(* IEC 61131-3 sources: llm-plc-st-eval/data/definitivo/claude-sonnet-4-6/B2/zero_shot, 3 files *)

(* ---- ejec_1.st ---- *)
```pascal
FUNCTION_BLOCK FB_Valvula
VAR_INPUT
    nivelAlto : BOOL; (* Sensor de nivel alto del tanque *)
END_VAR

VAR_OUTPUT
    valvula : BOOL; (* TRUE = válvula abierta, FALSE = válvula cerrada *)
END_VAR

VAR
    tonRetardo : TON; (* Temporizador de retardo para confirmación de nivel alto *)
END_VAR

(*
    Control de válvula de drenaje:
    - La válvula abre cuando nivelAlto permanece activo durante 5 segundos continuos.
    - La válvula cierra de inmediato si nivelAlto deja de estar activo.
*)

(* Activar temporizador solo mientras nivelAlto esté activo *)
tonRetardo(IN := nivelAlto, PT := T#5S);

(* La válvula abre cuando el temporizador completa los 5 segundos *)
(* Si nivelAlto cae, tonRetardo.Q se resetea de inmediato y la válvula cierra *)
valvula := tonRetardo.Q;

END_FUNCTION_BLOCK
```

(* ---- ejec_2.st ---- *)
```pascal
FUNCTION_BLOCK FB_Valvula
VAR_INPUT
    nivelAlto : BOOL; (* Sensor de nivel alto del tanque *)
END_VAR

VAR_OUTPUT
    valvula : BOOL; (* TRUE = válvula abierta, FALSE = válvula cerrada *)
END_VAR

VAR
    tonRetardo : TON; (* Temporizador de retardo para confirmar nivel alto *)
END_VAR

(*
    Control de válvula de drenaje:
    - La válvula abre cuando nivelAlto permanece activo durante 5 segundos continuos.
    - La válvula cierra de inmediato si nivelAlto deja de estar activo.
*)

(* Activar temporizador solo mientras nivelAlto esté activo *)
tonRetardo(IN := nivelAlto, PT := T#5S);

(* La válvula abre cuando el temporizador completa los 5 segundos *)
(* Si nivelAlto cae, tonRetardo.Q se pone FALSE de inmediato (IN=FALSE resetea el TON) *)
valvula := tonRetardo.Q;

END_FUNCTION_BLOCK
```

(* ---- ejec_3.st ---- *)
```pascal
FUNCTION_BLOCK FB_Valvula
VAR_INPUT
    nivelAlto : BOOL; (* Sensor de nivel alto del tanque *)
END_VAR

VAR_OUTPUT
    valvula : BOOL; (* TRUE = válvula abierta, FALSE = válvula cerrada *)
END_VAR

VAR
    tonRetardo : TON; (* Temporizador de retardo para confirmar nivel alto *)
END_VAR

(* ---------------------------------------------------------------
   Lógica de control:
   - El temporizador TON se habilita mientras nivelAlto esté activo.
   - Si nivelAlto se desactiva antes de 5 s, el temporizador se
     reinicia automáticamente (IN := FALSE).
   - Cuando nivelAlto permanece activo >= 5 s, tonRetardo.Q = TRUE
     y la válvula abre.
   - Si nivelAlto cae, la válvula cierra de inmediato (sin retardo).
--------------------------------------------------------------- *)

(* Llamada al temporizador: activo solo mientras nivelAlto sea TRUE *)
tonRetardo(
    IN := nivelAlto,
    PT := T#5S
);

(* La válvula abre cuando el temporizador confirma 5 s continuos de nivel alto.
   Si nivelAlto cae, tonRetardo.Q vuelve a FALSE de inmediato porque
   el temporizador se reinicia, cerrando la válvula sin retardo. *)
valvula := tonRetardo.Q;
```
